// TwinCAT 3 PLC project EventLoggerDemoPlc
// ProgramVersion: 3.1.4026.27
// libraries:
//   Tc2_Standard, * (Beckhoff Automation GmbH)
//   Tc2_System, * (Beckhoff Automation GmbH)
//   Tc3_EventLogger, * (Beckhoff Automation GmbH)
//   Tc3_Module, * (Beckhoff Automation GmbH)
// project tree:
//   DUTs/ E_HmiRequest.TcDUT, ST_HmiCommands.TcDUT, ST_HmiStatus.TcDUT, ST_PlcAlarm.TcDUT, ST_PlcAlarmTable.TcDUT
//   GVLs/ GVL_EventLogging.TcGVL, GVL_Hmi.TcGVL
//   POUs/Demo/ DemoMachine.TcPOU
//   POUs/EventLogging/ AlarmListener.TcPOU, AlarmPoint.TcPOU, MessagePoint.TcPOU
//   / PlcTask.TcTTO
//   POUs/ MAIN.TcPOU
// real-time tasks:
//   TASK PlcTask: cycle T#10ms, priority 20, ADS port 350

CONFIGURATION EventLoggerDemoPlc
    RESOURCE PLC ON TwinCAT3
        TASK PlcTask(INTERVAL := T#10ms, PRIORITY := 20);
        PROGRAM MAIN WITH PlcTask : MAIN;
    END_RESOURCE
END_CONFIGURATION

// ---- DUTs/E_HmiRequest.TcDUT
// Requests the HMI can make. Values are part of the HMI contract: never renumber.
{attribute 'qualified_only'}
{attribute 'strict'}
{attribute 'to_string'}
TYPE E_HmiRequest :
(
    NotSet              := 0,
    RaiseLowAirPressure := 1,
    ClearLowAirPressure := 2,
    RaiseDriveFault     := 3,
    ClearDriveFault     := 4,
    SendMachineStarted  := 5,
    SendBatchCompleted  := 6
) UINT;
END_TYPE

// ---- DUTs/ST_HmiCommands.TcDUT
// Written by the HMI. The HMI writes the arguments first and Request last.
// The PLC executes the request, increments Status.RequestCount and sets Request back to NotSet.
TYPE ST_HmiCommands :
STRUCT
    Request               : E_HmiRequest;
    IntegerArgument       : DINT;       // air pressure in mbar, drive error code, batch number
    SecondIntegerArgument : DINT;       // part count
    TextArgument          : STRING;     // operator name
    OvenTemperature       : LREAL := 20.0; // simulated process value, written by the HMI slider
END_STRUCT
END_TYPE

// ---- DUTs/ST_HmiStatus.TcDUT
// Read by the HMI.
TYPE ST_HmiStatus :
STRUCT
    Heartbeat             : UDINT;  // increments every cycle
    IsInitialised         : BOOL;   // all alarms and messages created in the EventLogger
    LastRequest           : E_HmiRequest;
    LastRequestAccepted   : BOOL;
    RequestCount          : UDINT;  // increments once per executed request
    OvenTemperature       : LREAL;
    OvenTemperatureLimit  : LREAL;
    OverTemperatureRaised : BOOL;
    LowAirPressureRaised  : BOOL;
    DriveFaultRaised      : BOOL;
END_STRUCT
END_TYPE

// ---- DUTs/ST_PlcAlarm.TcDUT
// One raised alarm, as reported to the PLC by the EventLogger.
TYPE ST_PlcAlarm :
STRUCT
    Entry         : TcEventEntry;   // event class GUID, event ID, severity
    SourceName    : STRING(80);
    TimeRaised    : ULINT;          // 100 ns since 1601-01-01 UTC (FILETIME)
    IsConfirmed   : BOOL;
    TextAvailable : BOOL;           // TRUE once the text has arrived, a few cycles after the raise
    Text          : T_MaxString;
END_STRUCT
END_TYPE

// ---- DUTs/ST_PlcAlarmTable.TcDUT
// Every alarm currently raised on this TwinCAT system, from any PLC or module.
TYPE ST_PlcAlarmTable :
STRUCT
    IsSubscribed : BOOL;
    Count        : UDINT;   // rows 0 to Count - 1 are in use, newest last
    Overflow     : BOOL;    // TRUE once an alarm could not be added because the table was full
    Alarms       : ARRAY[0..GVL_EventLogging.MaxPlcAlarms - 1] OF ST_PlcAlarm;
END_STRUCT
END_TYPE

// ---- GVLs/GVL_EventLogging.TcGVL
// Settings of the PLC-side alarm table.
{attribute 'qualified_only'}
VAR_GLOBAL CONSTANT
    MaxPlcAlarms         : UDINT := 32;     // rows in ST_PlcAlarmTable
    TextLanguageId       : DINT  := 1033;   // language of PLC-side texts, as a Windows LCID
    SubscribeRetryCycles : UDINT := 100;    // cycles between subscription attempts
END_VAR

// ---- GVLs/GVL_Hmi.TcGVL
// The HMI contract. The web HMI reads and writes these symbols by name over ADS.
{attribute 'qualified_only'}
VAR_GLOBAL
    Commands : ST_HmiCommands;
    Status   : ST_HmiStatus;
    PlcAlarms : ST_PlcAlarmTable;   // kept by AlarmListener from the EventLogger
END_VAR

// ---- POUs/MAIN.TcPOU
PROGRAM MAIN
VAR
    Machine  : DemoMachine;
    Listener : AlarmListener;
END_VAR

Machine.CyclicLogic(Commands := GVL_Hmi.Commands, Status := GVL_Hmi.Status);
Listener.CyclicLogic(Table := GVL_Hmi.PlcAlarms);

END_PROGRAM

// ---- POUs/Demo/DemoMachine.TcPOU
// The demo application. Supervises a simulated oven temperature and executes HMI requests,
// reporting everything through the TwinCAT EventLogger.
FUNCTION_BLOCK DemoMachine
VAR
    _OverTemperature : AlarmPoint;
    _LowAirPressure  : AlarmPoint;
    _DriveFault      : AlarmPoint;
    _MachineStarted  : MessagePoint;
    _BatchCompleted  : MessagePoint;
    _IsInitialised   : BOOL;
END_VAR
VAR CONSTANT
    OvenTemperatureLimit      : LREAL := 80.0;
    OvenTemperatureHysteresis : LREAL := 5.0;
END_VAR

METHOD CyclicLogic
VAR_IN_OUT
    Commands : ST_HmiCommands;
    Status   : ST_HmiStatus;
END_VAR
Status.Heartbeat := Status.Heartbeat + 1;

IF NOT _IsInitialised THEN
    _IsInitialised := Initialise();
END_IF
Status.IsInitialised := _IsInitialised;

IF NOT _IsInitialised THEN
    RETURN;
END_IF

SuperviseOvenTemperature(Temperature := Commands.OvenTemperature);

IF Commands.Request <> E_HmiRequest.NotSet THEN
    Status.LastRequest         := Commands.Request;
    Status.LastRequestAccepted := HandleRequest(Commands := Commands);
    Status.RequestCount        := Status.RequestCount + 1;
    Commands.Request           := E_HmiRequest.NotSet;
END_IF

Status.OvenTemperature       := Commands.OvenTemperature;
Status.OvenTemperatureLimit  := OvenTemperatureLimit;
Status.OverTemperatureRaised := _OverTemperature.IsRaised;
Status.LowAirPressureRaised  := _LowAirPressure.IsRaised;
Status.DriveFaultRaised      := _DriveFault.IsRaised;
END_METHOD

METHOD PRIVATE Initialise : BOOL
// Creates every alarm and message. Safe to call again after a partial failure.
VAR
    AlarmsCreated   : BOOL;
    MessagesCreated : BOOL;
END_VAR
// AND does not short-circuit, so every Create is attempted on every call.
AlarmsCreated := _OverTemperature.Create(Entry := TC_EVENTS.EventLoggerDemo.OverTemperature, WithConfirmation := TRUE, SourceName := 'Oven')
             AND _LowAirPressure.Create(Entry := TC_EVENTS.EventLoggerDemo.LowAirPressure, WithConfirmation := FALSE, SourceName := 'Air supply')
             AND _DriveFault.Create(Entry := TC_EVENTS.EventLoggerDemo.DriveFault, WithConfirmation := TRUE, SourceName := 'Conveyor drive');

MessagesCreated := _MachineStarted.Create(Entry := TC_EVENTS.EventLoggerDemo.MachineStarted, SourceName := 'Operator panel')
               AND _BatchCompleted.Create(Entry := TC_EVENTS.EventLoggerDemo.BatchCompleted, SourceName := 'Production');

Initialise := AlarmsCreated AND MessagesCreated;
END_METHOD

METHOD PRIVATE SuperviseOvenTemperature
// Raises OverTemperature above the limit and clears it below limit minus hysteresis.
VAR_INPUT
    Temperature : LREAL;
END_VAR
IF NOT _OverTemperature.IsRaised THEN
    IF Temperature > OvenTemperatureLimit THEN
        _OverTemperature.NewArguments().AddDINT(LREAL_TO_DINT(Temperature)).AddDINT(LREAL_TO_DINT(OvenTemperatureLimit));
        _OverTemperature.Raise();
    END_IF
ELSIF Temperature < OvenTemperatureLimit - OvenTemperatureHysteresis THEN
    _OverTemperature.Clear(ResetConfirmation := FALSE);
END_IF
END_METHOD

METHOD PRIVATE HandleRequest : BOOL
// Executes one HMI request. Returns TRUE if the EventLogger accepted it.
VAR_IN_OUT CONSTANT
    Commands : ST_HmiCommands;
END_VAR
CASE Commands.Request OF
    E_HmiRequest.RaiseLowAirPressure:
        IF _LowAirPressure.IsRaised THEN
            HandleRequest := TRUE;
        ELSE
            _LowAirPressure.NewArguments().AddDINT(Commands.IntegerArgument);
            HandleRequest := _LowAirPressure.Raise();
        END_IF

    E_HmiRequest.ClearLowAirPressure:
        HandleRequest := _LowAirPressure.Clear(ResetConfirmation := FALSE);

    E_HmiRequest.RaiseDriveFault:
        IF _DriveFault.IsRaised THEN
            HandleRequest := TRUE;
        ELSE
            _DriveFault.NewArguments().AddDINT(Commands.IntegerArgument);
            HandleRequest := _DriveFault.Raise();
        END_IF

    E_HmiRequest.ClearDriveFault:
        // Clearing does not confirm: the alarm stays in the list until the operator confirms it.
        HandleRequest := _DriveFault.Clear(ResetConfirmation := FALSE);

    E_HmiRequest.SendMachineStarted:
        _MachineStarted.NewArguments().AddString(Commands.TextArgument);
        HandleRequest := _MachineStarted.Send();

    E_HmiRequest.SendBatchCompleted:
        _BatchCompleted.NewArguments().AddDINT(Commands.IntegerArgument).AddDINT(Commands.SecondIntegerArgument);
        HandleRequest := _BatchCompleted.Send();

ELSE
    HandleRequest := FALSE;
END_CASE
END_METHOD

END_FUNCTION_BLOCK

// ---- POUs/EventLogging/AlarmPoint.TcPOU
// One alarm in the TwinCAT EventLogger, with its own source name.
// Call Create once before anything else. Fill arguments with NewArguments() before Raise.
FUNCTION_BLOCK AlarmPoint
VAR
    _Alarm      : FB_TcAlarm;
    _Source     : FB_TcSourceInfo;
    _IsCreated  : BOOL;
    _LastResult : HRESULT;
END_VAR

METHOD Create : BOOL
// Creates the alarm instance in the EventLogger. Returns TRUE at once if already created.
VAR_INPUT
    Entry            : TcEventEntry;   // e.g. TC_EVENTS.EventLoggerDemo.OverTemperature
    WithConfirmation : BOOL;
    SourceName       : STRING;         // shown as the alarm's source
END_VAR
IF _IsCreated THEN
    Create := TRUE;
    RETURN;
END_IF

_Source.Clear();
_Source.sName := SourceName;

_LastResult := _Alarm.CreateEx(stEventEntry := Entry, bWithConfirmation := WithConfirmation, ipSourceInfo := _Source);
_IsCreated := (_LastResult >= 0);
Create := _IsCreated;
END_METHOD

METHOD NewArguments : I_TcArguments
// Empties the argument list and returns it for chaining: NewArguments().AddDINT(42).AddDINT(7)
// Arguments are captured when the alarm is raised.
NewArguments := _Alarm.ipArguments.Clear();
END_METHOD

METHOD Raise : BOOL
IF NOT _IsCreated THEN
    Raise := FALSE;
    RETURN;
END_IF

_LastResult := _Alarm.Raise(nTimeStamp := 0);
Raise := (_LastResult >= 0);
END_METHOD

METHOD Clear : BOOL
VAR_INPUT
    ResetConfirmation : BOOL;   // TRUE: an unconfirmed alarm can no longer be confirmed
END_VAR
IF NOT _IsCreated THEN
    Clear := FALSE;
    RETURN;
END_IF

_LastResult := _Alarm.Clear(nTimeStamp := 0, bResetConfirmation := ResetConfirmation);
Clear := (_LastResult >= 0);
END_METHOD

PROPERTY IsCreated : BOOL
GET
IsCreated := _IsCreated;
END_GET
END_PROPERTY

PROPERTY IsRaised : BOOL
GET
IsRaised := _IsCreated AND_THEN _Alarm.bRaised;
END_GET
END_PROPERTY

PROPERTY LastResult : HRESULT
GET
LastResult := _LastResult;
END_GET
END_PROPERTY

END_FUNCTION_BLOCK

// ---- POUs/EventLogging/MessagePoint.TcPOU
// One message in the TwinCAT EventLogger, with its own source name.
// Call Create once before anything else. Fill arguments with NewArguments() before Send.
FUNCTION_BLOCK MessagePoint
VAR
    _Message    : FB_TcMessage;
    _Source     : FB_TcSourceInfo;
    _IsCreated  : BOOL;
    _LastResult : HRESULT;
END_VAR

METHOD Create : BOOL
// Creates the message instance in the EventLogger. Returns TRUE at once if already created.
VAR_INPUT
    Entry      : TcEventEntry;   // e.g. TC_EVENTS.EventLoggerDemo.MachineStarted
    SourceName : STRING;         // shown as the message's source
END_VAR
IF _IsCreated THEN
    Create := TRUE;
    RETURN;
END_IF

_Source.Clear();
_Source.sName := SourceName;

_LastResult := _Message.CreateEx(stEventEntry := Entry, ipSourceInfo := _Source);
_IsCreated := (_LastResult >= 0);
Create := _IsCreated;
END_METHOD

METHOD NewArguments : I_TcArguments
// Empties the argument list and returns it for chaining: NewArguments().AddString(Name)
NewArguments := _Message.ipArguments.Clear();
END_METHOD

METHOD Send : BOOL
IF NOT _IsCreated THEN
    Send := FALSE;
    RETURN;
END_IF

_LastResult := _Message.Send(nTimeStamp := 0);
Send := (_LastResult >= 0);
END_METHOD

PROPERTY IsCreated : BOOL
GET
IsCreated := _IsCreated;
END_GET
END_PROPERTY

PROPERTY LastResult : HRESULT
GET
LastResult := _LastResult;
END_GET
END_PROPERTY

END_FUNCTION_BLOCK

// ---- POUs/EventLogging/AlarmListener.TcPOU
// Keeps a table of the alarms currently raised on this TwinCAT system, by listening to the
// EventLogger. Call CyclicLogic every cycle; the table it is given is updated during the call.
FUNCTION_BLOCK AlarmListener EXTENDS FB_ListenerBase2
VAR
    _Table           : REFERENCE TO ST_PlcAlarmTable;
    _IsSubscribed    : BOOL;
    _SubscribeResult : HRESULT;
    _ExecuteResult   : HRESULT;
    _RetryCountdown  : UDINT;

    // Alarm texts arrive asynchronously, a few cycles after the alarm is raised. One request
    // slot per possible row; a slot is matched back to its row by event and source, because
    // rows move when others are removed.
    _TextRequests : ARRAY[0..GVL_EventLogging.MaxPlcAlarms - 1] OF FB_RequestEventText;
    _TextPending  : ARRAY[0..GVL_EventLogging.MaxPlcAlarms - 1] OF BOOL;
    _TextDiscard  : ARRAY[0..GVL_EventLogging.MaxPlcAlarms - 1] OF BOOL;
    _TextEntry    : ARRAY[0..GVL_EventLogging.MaxPlcAlarms - 1] OF TcEventEntry;
    _TextSource   : ARRAY[0..GVL_EventLogging.MaxPlcAlarms - 1] OF STRING(80);
END_VAR

METHOD PRIVATE CollectTexts
// Copies each finished text into its alarm's row. A row removed in the meantime is skipped.
VAR
    Slot : DINT;
    Row  : DINT;
END_VAR
FOR Slot := 0 TO UDINT_TO_DINT(GVL_EventLogging.MaxPlcAlarms) - 1 DO
    IF NOT _TextPending[Slot] OR_ELSE _TextRequests[Slot].bBusy THEN
        CONTINUE;
    END_IF

    _TextPending[Slot] := FALSE;
    IF _TextDiscard[Slot] OR_ELSE _TextRequests[Slot].bError THEN
        CONTINUE;
    END_IF

    Row := FindAlarm(Entry := _TextEntry[Slot], SourceName := _TextSource[Slot]);
    IF Row >= 0 THEN
        _TextRequests[Slot].GetString(sResult := _Table.Alarms[Row].Text, nResult := SIZEOF(_Table.Alarms[Row].Text));
        _Table.Alarms[Row].TextAvailable := TRUE;
    END_IF
END_FOR
END_METHOD

METHOD CyclicLogic
// Subscribes on first use, then processes the EventLogger's queue. Callbacks run inside Execute,
// so Table is valid whenever they write to it.
VAR_IN_OUT
    Table : ST_PlcAlarmTable;
END_VAR
_Table REF= Table;

IF NOT _IsSubscribed THEN
    IF _RetryCountdown > 0 THEN
        _RetryCountdown := _RetryCountdown - 1;
    ELSE
        _SubscribeResult := THIS^.Subscribe(ipMessageFilterConfig := 0, ipAlarmFilterConfig := 0);
        _IsSubscribed := (_SubscribeResult >= 0);
        _RetryCountdown := GVL_EventLogging.SubscribeRetryCycles;
    END_IF
END_IF

Table.IsSubscribed := _IsSubscribed;

IF _IsSubscribed THEN
    _ExecuteResult := THIS^.Execute();
END_IF

CollectTexts();
END_METHOD

PROPERTY ExecuteResult : HRESULT
GET
ExecuteResult := _ExecuteResult;
END_GET
END_PROPERTY

METHOD PRIVATE FindAlarm : DINT
// Returns the row of the alarm with this event class, event ID and source, or -1.
VAR_INPUT
    Entry      : TcEventEntry;
    SourceName : STRING(80);
END_VAR
VAR
    Row : DINT;
END_VAR
FindAlarm := -1;
FOR Row := 0 TO UDINT_TO_DINT(_Table.Count) - 1 DO
    IF IsSameAlarm(EntryA := _Table.Alarms[Row].Entry, SourceA := _Table.Alarms[Row].SourceName, EntryB := Entry, SourceB := SourceName) THEN
        FindAlarm := Row;
        RETURN;
    END_IF
END_FOR
END_METHOD

METHOD PRIVATE IsSameAlarm : BOOL
// The EventLogger tells alarms apart by event class, event ID and source.
VAR_INPUT
    EntryA  : TcEventEntry;
    SourceA : STRING(80);
    EntryB  : TcEventEntry;
    SourceB : STRING(80);
END_VAR
IsSameAlarm := MEMCMP(ADR(EntryA.uuidEventClass), ADR(EntryB.uuidEventClass), SIZEOF(GUID)) = 0
               AND_THEN EntryA.nEventId = EntryB.nEventId
               AND_THEN SourceA = SourceB;
END_METHOD

PROPERTY IsSubscribed : BOOL
GET
IsSubscribed := _IsSubscribed;
END_GET
END_PROPERTY

METHOD OnAlarmCleared : HRESULT
VAR_INPUT
    fbEvent : REFERENCE TO FB_TcEvent;
END_VAR
VAR
    Entry      : TcEventEntry;
    SourceName : STRING(80);
    Index      : DINT;
END_VAR
// The table lists raised alarms only, so a cleared alarm leaves it, confirmed or not.
OnAlarmCleared := 0;
IF NOT __ISVALIDREF(_Table) THEN
    RETURN;
END_IF

Entry := fbEvent.stEventEntry;
SourceName := SourceNameOf(fbEvent := fbEvent);
Index := FindAlarm(Entry := Entry, SourceName := SourceName);
IF Index >= 0 THEN
    RemoveAt(Index := Index);
END_IF
END_METHOD

METHOD OnAlarmConfirmed : HRESULT
VAR_INPUT
    fbEvent : REFERENCE TO FB_TcEvent;
END_VAR
VAR
    Entry      : TcEventEntry;
    SourceName : STRING(80);
    Index      : DINT;
END_VAR
OnAlarmConfirmed := 0;
IF NOT __ISVALIDREF(_Table) THEN
    RETURN;
END_IF

Entry := fbEvent.stEventEntry;
SourceName := SourceNameOf(fbEvent := fbEvent);
Index := FindAlarm(Entry := Entry, SourceName := SourceName);
IF Index >= 0 THEN
    _Table.Alarms[Index].IsConfirmed := TRUE;
END_IF
END_METHOD

METHOD OnAlarmDisposed : HRESULT
VAR_INPUT
    fbEvent : REFERENCE TO FB_TcEvent;
END_VAR
VAR
    Entry      : TcEventEntry;
    SourceName : STRING(80);
    Index      : DINT;
END_VAR
// The alarm instance was released, for example because its PLC stopped.
OnAlarmDisposed := 0;
IF NOT __ISVALIDREF(_Table) THEN
    RETURN;
END_IF

Entry := fbEvent.stEventEntry;
SourceName := SourceNameOf(fbEvent := fbEvent);
Index := FindAlarm(Entry := Entry, SourceName := SourceName);
IF Index >= 0 THEN
    RemoveAt(Index := Index);
END_IF
END_METHOD

METHOD OnAlarmRaised : HRESULT
VAR_INPUT
    fbEvent : REFERENCE TO FB_TcEvent;
END_VAR
VAR
    Entry      : TcEventEntry;
    SourceName : STRING(80);
    Index      : DINT;
END_VAR
OnAlarmRaised := 0;
IF NOT __ISVALIDREF(_Table) THEN
    RETURN;
END_IF

Entry := fbEvent.stEventEntry;
SourceName := SourceNameOf(fbEvent := fbEvent);

Index := FindAlarm(Entry := Entry, SourceName := SourceName);
IF Index < 0 THEN
    IF _Table.Count >= GVL_EventLogging.MaxPlcAlarms THEN
        _Table.Overflow := TRUE;
        RETURN;
    END_IF
    Index := UDINT_TO_DINT(_Table.Count);
    _Table.Count := _Table.Count + 1;
END_IF

_Table.Alarms[Index].Entry       := Entry;
_Table.Alarms[Index].SourceName  := SourceName;
_Table.Alarms[Index].TimeRaised  := fbEvent.nTimestamp;
_Table.Alarms[Index].IsConfirmed := FALSE;
_Table.Alarms[Index].TextAvailable := FALSE;
_Table.Alarms[Index].Text := '';
StartTextRequest(fbEvent := fbEvent, Entry := Entry, SourceName := SourceName);
END_METHOD

METHOD PRIVATE RemoveAt
// Removes one row and closes the gap, keeping the remaining rows in order.
VAR_INPUT
    Index : DINT;
END_VAR
VAR
    Row   : DINT;
    Empty : ST_PlcAlarm;
END_VAR
IF Index < 0 OR_ELSE Index >= UDINT_TO_DINT(_Table.Count) THEN
    RETURN;
END_IF

FOR Row := Index TO UDINT_TO_DINT(_Table.Count) - 2 DO
    _Table.Alarms[Row] := _Table.Alarms[Row + 1];
END_FOR

_Table.Count := _Table.Count - 1;
_Table.Alarms[_Table.Count] := Empty;
END_METHOD

METHOD PRIVATE SourceNameOf : STRING(80)
VAR_INPUT
    fbEvent : REFERENCE TO FB_TcEvent;
END_VAR
IF fbEvent.ipSourceInfo <> 0 THEN
    SourceNameOf := fbEvent.ipSourceInfo.sName;
ELSE
    SourceNameOf := '';
END_IF
END_METHOD

METHOD PRIVATE StartTextRequest
// Starts the asynchronous text request for a raised alarm. Called inside the callback, while
// fbEvent and its arguments are valid; CollectTexts picks the text up when it arrives.
VAR_INPUT
    fbEvent    : REFERENCE TO FB_TcEvent;
    Entry      : TcEventEntry;
    SourceName : STRING(80);
END_VAR
VAR
    Slot     : DINT;
    FreeSlot : DINT;
END_VAR
FreeSlot := -1;
FOR Slot := 0 TO UDINT_TO_DINT(GVL_EventLogging.MaxPlcAlarms) - 1 DO
    IF _TextPending[Slot] THEN
        // A request still running for the same alarm belongs to an earlier raise.
        IF IsSameAlarm(EntryA := _TextEntry[Slot], SourceA := _TextSource[Slot], EntryB := Entry, SourceB := SourceName) THEN
            _TextDiscard[Slot] := TRUE;
        END_IF
    ELSIF FreeSlot < 0 THEN
        FreeSlot := Slot;
    END_IF
END_FOR

IF FreeSlot < 0 THEN
    RETURN; // every slot busy: this row keeps TextAvailable FALSE
END_IF

_TextEntry[FreeSlot]   := Entry;
_TextSource[FreeSlot]  := SourceName;
_TextDiscard[FreeSlot] := FALSE;
_TextPending[FreeSlot] := TRUE;
_TextRequests[FreeSlot].Request(eventClass := Entry.uuidEventClass, nEventId := Entry.nEventId, nLangId := GVL_EventLogging.TextLanguageId, ipArgs := fbEvent.ipArguments);
END_METHOD

PROPERTY SubscribeResult : HRESULT
GET
SubscribeResult := _SubscribeResult;
END_GET
END_PROPERTY

END_FUNCTION_BLOCK
